Fanuc KAREL source: KD00075.KL

PROGRAM KD00075
%NOLOCKGROUP
VAR
  I: INTEGER
  J: INTEGER
  B: BOOLEAN
  R: REAL
  S: STRING[80]
BEGIN
  CONDITION[1]:
  WHEN DIN[1] = ON DO
    I = 1
  ENDCONDITION
END KD00075
